(* IEC 61131-3 sources: model-first-plc-agent-ai/results/T2-B-30, 1 file *)

(* ---- b_code.st ---- *)
FUNCTION_BLOCK FillingControl
VAR_INPUT
    start : BOOL;
    stop : BOOL;
    LSH : BOOL;
    LSHH : BOOL;
    TimerDuration : TIME;
END_VAR
VAR_OUTPUT
    fill_valve : BOOL;
    discharge_valve : BOOL;
END_VAR
VAR
    current_state : INT := 0;
    filling_timer : TON;
    timer_done : BOOL := FALSE;
END_VAR

IF stop THEN
    current_state := 0;
ELSE
    CASE current_state OF
        0:
            IF start AND NOT LSHH THEN
                current_state := 1;
            END_IF;
        1:
            current_state := 1;
    ELSE
        current_state := 0;
    END_CASE;
END_IF;

filling_timer(
    IN := (current_state = 1) AND NOT stop AND NOT LSHH,
    PT := TimerDuration
);
timer_done := filling_timer.Q;

IF (current_state = 1) AND (timer_done OR LSHH) THEN
    current_state := 0;
END_IF;

fill_valve := (current_state = 1) AND NOT stop AND NOT LSHH;
discharge_valve := FALSE;

(* Reset immediately so a new start on the next scan gets a fresh timer. *)
IF current_state = 0 THEN
    filling_timer(IN := FALSE, PT := TimerDuration);
    timer_done := filling_timer.Q;
END_IF;

END_FUNCTION_BLOCK

PROGRAM Main
VAR
    StartCommand AT %IX100.0 : BOOL;
    StopCommand AT %IX100.1 : BOOL;
    LSH AT %IX100.2 : BOOL;
    LSHH AT %IX100.3 : BOOL;
    FillValve AT %QX100.0 : BOOL;
    DischargeValve AT %QX100.1 : BOOL;
END_VAR
VAR
    TimerDuration : TIME := T#10s;
    start_edge : R_TRIG;
    controller : FillingControl;
END_VAR

start_edge(CLK := StartCommand);

controller(
    start := start_edge.Q,
    stop := StopCommand,
    LSH := LSH,
    LSHH := LSHH,
    TimerDuration := TimerDuration
);

FillValve := controller.fill_valve;
DischargeValve := controller.discharge_valve;

END_PROGRAM
